FUNCTION_BLOCK FB_MotorSim EXTENDS FB_MotorBase

(* Base bodies run only when called explicitly. Shared Update is inherited. *)
SUPER^();

END_FUNCTION_BLOCK

(* stored: Version 1.1.0.1, ProductVersion 3.1 *)
